Fanuc KAREL source: KT00891.KL

PROGRAM KT00891
%NOLOCKGROUP
VAR
  P1: JOINTPOS
  P2: JOINTPOS
  OUT: POSITION
BEGIN
  OUT = INV(P1)
END KT00891
